(* KBO mirror coating selector (Si/B4C) core, an abstract base by convention:
   thin ND-framework state-mover wrapper that holds only references, interfaces
   and fbStates. The state bridge is here as REFERENCE TO UINT (eEnumSetRef and
   eEnumGetRef) and the body runs on it, but the enum variables, the state
   storage and the state names belong to the derived type
   (FB_KBO_Coating_States), which passes them in.

   A derived type supplies everything that depends on the state list:
     - eEnumSet and eEnumGet, the device enum (UINT base, OUT = 1, then the
       targets) with the MMS:STATE:SET and MMS:STATE:GET pytmc pragmas, so the
       EPICS state menu comes from that enum;
     - afbStateDefaults, one FB_CC_InternalStateConfig per state, which writes
       the per-state sName and fDelta;
     - an FB_Init that repeats the inputs below and binds eEnumSetRef and
       eEnumGetRef to the enum variables, and a CallAfterInit that calls the
       configurators. The base CallAfterInit runs on its own through the
       call_after_init attribute.
   FB_KBO_Coating_States is the library derived type (E_KBO_CoatingStates).
*)
{attribute 'call_after_init'}
FUNCTION_BLOCK FB_KBO_Coating_States_Core
VAR
    {attribute 'no_copy'}
    aiMotionStage         : REFERENCE TO ARRAY[1..MotionConstants.MAX_STATE_MOTORS] OF I_MotionStage;
    {attribute 'no_copy'}
    astPositionState      : REFERENCE TO ARRAY[1..MotionConstants.MAX_STATE_MOTORS]
                                            OF ARRAY[1..GeneralConstants.MAX_STATES] OF ST_PositionState;
    {attribute 'no_copy'}
    fbFFHWO               : REFERENCE TO FB_HardwareFFOutput;
    {attribute 'no_copy'}
    fbArbiter             : REFERENCE TO FB_Arbiter;
    sDeviceName           : STRING;
    sTransitionKey        : STRING;
    bEnableMotion         : BOOL := TRUE;
    bEnableBeamParams     : BOOL;
    bEnablePositionLimits : BOOL;
    bReadDBNow            : BOOL;
    bFileReaderBusy       : REFERENCE TO BOOL;
    bFileReaderError      : REFERENCE TO BOOL;

    (* State bridge, bound by the derived type to its enum variables.
       eEnumSetRef receives move requests and eEnumGetRef reports the
       current state. Both are UINT views of those variables. *)
    {attribute 'no_copy'}
    eEnumSetRef           : REFERENCE TO UINT;
    {attribute 'no_copy'}
    eEnumGetRef           : REFERENCE TO UINT;

    {attribute 'pytmc' := 'pv: MMS'}
    fbStates : FB_PositionStatePMPSND(
        aiMotionStage         := aiMotionStage,
        astPositionState      := astPositionState,
        nActiveMotorCount     := nStateMotorCount,
        eEnumSet              := eEnumSetRef,
        eEnumGet              := eEnumGetRef,
        bEnableMotion         := bEnableMotion,
        eMotionRequestPolicy  := E_MotionRequestPolicy.INTERRUPT,
        bEnableBeamParams     := bEnableBeamParams,
        bEnablePositionLimits := bEnablePositionLimits,
        bReadDBNow            := bReadDBNow,
        bFileReaderBusy       := bFileReaderBusy,
        bFileReaderError      := bFileReaderError,
        fbFFHWO               := fbFFHWO,
        fbArbiter             := fbArbiter,
        sDeviceName           := sDeviceName,
        sTransitionKey        := sTransitionKey
    );
END_VAR
VAR_OUTPUT
    // The PMPS database lookup associated with the current position state.
    stDbStateParams: ST_DbStateParams;
END_VAR
VAR CONSTANT
    (* Number of motors the state mover drives. Every device here has one state
       motor, in slot 1; the code around fbStates assumes it. *)
    nStateMotorCount : UINT := 1;
    // State in-position tolerance, applied per-state by afbStateDefaults.
    // Units in Millimeters (matches prior install values).
    FDELTA_DEFAULT  : LREAL := 0.1;
    // Reference motion dynamics for this mirror - NOT applied by this FB.
    // The caller sets these on the motor (e.g. SetMotionParam) or relies
    // on the NC axis's own configured defaults. Y/X pair documents what
    // the prior install used, for whoever wires up a real axis.
    FVELOCITY_DEFAULT : LREAL := 0.150;
    FYACCEL_DEFAULT   : LREAL := 10;
    FYDECEL_DEFAULT   : LREAL := 10;
    FXACCEL_DEFAULT   : LREAL := 100;
    FXDECEL_DEFAULT   : LREAL := 100;
END_VAR

IF NOT __ISVALIDREF(aiMotionStage)
   OR NOT __ISVALIDREF(astPositionState)
   OR NOT __ISVALIDREF(fbFFHWO)
   OR NOT __ISVALIDREF(fbArbiter)
   OR NOT __ISVALIDREF(eEnumSetRef)
   OR NOT __ISVALIDREF(eEnumGetRef) THEN
    RETURN;
END_IF

fbStates(
    stDbStateParams => stDbStateParams
);

(* Auto-fired after FB_Init. Wires fbStates through CallAfterInitCore. *)
{attribute 'call_after_init'}
METHOD CallAfterInit
THIS^.CallAfterInitCore();
END_METHOD

(* Wires fbStates with the references this FB holds, through
   CallAfterInitStateMover / CallAfterInitPMPS, because fbStates' inline-init
   ran first and forwarded nil refs. Does nothing while the essential refs are
   still nil. CallAfterInit calls it. A derived type that was re-wired after its
   host FB's CallAfterInit calls it again through SUPER^. *)
METHOD CallAfterInitCore
IF NOT __ISVALIDREF(aiMotionStage)
   OR NOT __ISVALIDREF(astPositionState)
   OR NOT __ISVALIDREF(eEnumSetRef)
   OR NOT __ISVALIDREF(eEnumGetRef) THEN
    RETURN;
END_IF

THIS^.fbStates.CallAfterInitStateMover(
    aiMotionStage         := aiMotionStage,
    astPositionState      := astPositionState,
    nActiveMotorCount     := nStateMotorCount,
    eEnumSet              := eEnumSetRef,
    eEnumGet              := eEnumGetRef,
    bEnableMotion         := bEnableMotion,
    eMotionRequestPolicy  := E_MotionRequestPolicy.INTERRUPT,
);

THIS^.fbStates.CallAfterInitPMPS(
    aiMotionStage         := aiMotionStage,
    astPositionState      := astPositionState,
    bEnableBeamParams     := bEnableBeamParams,
    bEnablePositionLimits := bEnablePositionLimits,
    bReadDBNow            := bReadDBNow,
    bFileReaderBusy       := bFileReaderBusy,
    bFileReaderError      := bFileReaderError,
    fbFFHWO               := fbFFHWO,
    fbArbiter             := fbArbiter,
    sDeviceName           := sDeviceName,
    sTransitionKey        := sTransitionKey
);
END_METHOD

(* Stores FB_Init inputs into instance fields; every non-value input is
   REFERENCE TO, REF= bound for the FB lifetime. fbStates inline-init
   captured these params at construction, so this records the same refs
   on THIS^ for body use and live caller writes. *)
{attribute 'analysis' := '-33'}
METHOD FB_Init : BOOL
VAR_INPUT
    bInitRetains           : BOOL;
    bInCopyCode            : BOOL;
    aiMotionStage          : REFERENCE TO ARRAY[1..MotionConstants.MAX_STATE_MOTORS] OF I_MotionStage;
    astPositionState       : REFERENCE TO ARRAY[1..MotionConstants.MAX_STATE_MOTORS]
                                            OF ARRAY[1..GeneralConstants.MAX_STATES] OF ST_PositionState;
    fbFFHWO                : REFERENCE TO FB_HardwareFFOutput;
    fbArbiter              : REFERENCE TO FB_Arbiter;
    sDeviceName            : STRING;
    sTransitionKey         : STRING;
    bEnableBeamParams      : BOOL;
    bEnablePositionLimits  : BOOL;
    bReadDBNow             : BOOL;
    bFileReaderBusy        : REFERENCE TO BOOL;
    bFileReaderError       : REFERENCE TO BOOL;
END_VAR
THIS^.aiMotionStage    REF= aiMotionStage;
THIS^.astPositionState REF= astPositionState;
THIS^.fbFFHWO          REF= fbFFHWO;
THIS^.fbArbiter        REF= fbArbiter;
THIS^.sDeviceName      := sDeviceName;
THIS^.sTransitionKey   := sTransitionKey;
THIS^.bEnableBeamParams     := bEnableBeamParams;
THIS^.bEnablePositionLimits := bEnablePositionLimits;
THIS^.bReadDBNow            := bReadDBNow;
THIS^.bFileReaderBusy       REF= bFileReaderBusy;
THIS^.bFileReaderError      REF= bFileReaderError;
END_METHOD

END_FUNCTION_BLOCK

(* stored: Version 1.1.0.1
   POU FB_KBO_Coating_States_Core: Id {1bf9e26b-e907-4179-b0ff-e94e256de3ba}, SpecialFunc None
   Method CallAfterInit: Id {21a653fa-0b7a-4428-9b61-4f0f09b1e25d}
   Method CallAfterInitCore: Id {423a868f-985a-4282-84f1-a14056ccb609}
   Method FB_Init: Id {07fc869a-3706-4f0f-ac2f-6f69077c3bd7} *)
